// TIA Portal V20 export
// export: Created 2026-10-12T15:52:18.2848565Z, ExportSetting WithDefaults, DisplayName Totally Integrated Automation Portal, DisplayVersion V20, DisplayName TIA Portal Openness, DisplayVersion V20, DisplayName TIA Portal Teamcenter Gateway, DisplayVersion V20, DisplayName TIA Portal Version Control Interface, DisplayVersion V20, DisplayName SINAMICS Startdrive Advanced, DisplayVersion V20 SP1 Update 2, DisplayName SINAMICS Startdrive G110M, G120, G120C, G120D, G120P, G115D, DisplayVersion V20 SP1 Update 2, DisplayName SINAMICS Startdrive G130, G150, S120, S150, SINAMICS MV, G220, S200, S210, DisplayVersion V20 SP1 Update 2, DisplayName STEP 7 Professional, DisplayVersion V20, DisplayName STEP 7 Safety, DisplayVersion V20, DisplayName WinCC Basic/Comfort/Advanced, DisplayVersion V20, DisplayName WinCC Professional, DisplayVersion V20, DisplayName WinCC Unified, DisplayVersion V20
FUNCTION "FRK_AlarmHistoryHeaderSave" : Void   // FC43, SCL
{ S7_Optimized_Access := 'TRUE' }
VERSION : 0.1
// stored: AutoNumber true, IsIECCheckEnabled false, SetENOAutomatically false, UDAEnableTagReadback false
   VAR_IN_OUT
      AlarmLog : "FRK_AlarmLog";
   END_VAR
   VAR_TEMP
      Slot : Int;
   END_VAR
BEGIN

   #Slot := #AlarmLog.HistorySlot;
   IF #Slot < 1 OR #Slot > 3 THEN
       RETURN;
   END_IF;
   "FRK_AlarmHistory".Rows[#Slot].SchemaVersion := 1;
   "FRK_AlarmHistory".Rows[#Slot].Generation := "FRK_AccessNext"(Previous := "FRK_AlarmHistory".Rows[#Slot].Generation);
   "FRK_AlarmHistory".Rows[#Slot].RingHead := #AlarmLog.RingHead;
   "FRK_AlarmHistory".Rows[#Slot].RingUsed := #AlarmLog.RingUsed;
   "FRK_AlarmHistory".Rows[#Slot].Truncated := #AlarmLog.Truncated;
   "FRK_AlarmHistory".Rows[#Slot].Checksum := "FRK_AlarmHistoryHeaderCrc"(Slot := #Slot);
   "FRK_AlarmHistory".Commissioned[#Slot] := TRUE;
END_FUNCTION
